Fanuc KAREL source: KT00455.KL

PROGRAM KT00455
%NOLOCKGROUP
VAR
  P1: POSITION
  P2: POSITION
  OUT: BOOLEAN
BEGIN
  OUT = P1 >= P2
END KT00455
